(* IEC 61131-3 sources: SortJet_MasterSPS_Aufbau.fbsproj/09_Station/Stationen/Anlegetisch[201,205]/Aktionen, 2 files *)

(* ---- Anlegetisch_Austransport_FB_V01_00_00.fb.st ---- *)
(* METADATA
{
	"v3Meta": {
		"objectGuid": "29c6a30c-ea89-4d6e-bcb0-e2d154ff9fe9"
	}
}
*)
FUNCTION_BLOCK Anlegetisch_Austransport_FB_V01_00_00 EXTENDS Basic_Station_Austransport_FB_V01_00_00
(* Hinweis:
   - Austransport des Anlegetisches: Hubrahmen ausfahren, Austransport, Hubrahmen absenken, sobald die Sensorik
     frei ist, danach die Achsen des Glastransports abnullen
   - Der Rumpf ersetzt den Rumpf des Basic-Austransports, die Komponenten (Glastransport) kommen vom Basic-Baustein
*)
VAR_INPUT

  // Bausteine
  Hubrahmen : REFERENCE TO ZylinderPneumatik_Riemen_FB_V01_00_00;

END_VAR
//-------------------------------------------------------------------------------------------------
// AKTION: AUSTRANSPORT
//-------------------------------------------------------------------------------------------------
IF ( BasisStationsParameter.bAustransport[wWand]
     AND bpAutomatikAktiv )
THEN

  // Ausnahmesituation
  IF ( Glastransport.bpFehler ) THEN
    Glastransport.bpAustransport := FALSE;
    Glastransport.bpReferenz     := FALSE;
    BasisStationsParameter.wFehlerNummer := Glastransport.wpFehlerNr;
    steplAktion := STEP_900_E;
  END_IF

  IF ( Hubrahmen.bpFehler ) THEN
    Hubrahmen.bpStartAusfahren := FALSE;
    BasisStationsParameter.awFehlerInformationen[1] := cZYLINDER_HUBRAHMEN;
    BasisStationsParameter.wFehlerNummer := Hubrahmen.wpFehlerNr;
    steplAktion := STEP_900_E;
  END_IF

  CASE steplAktion OF
    // AUSTRANSPORT ==============================
    STEP_0_E:
      (* Hinweis:
         - -
      *)
      bpFehler := FALSE;
      Hubrahmen.bpStartAusfahren := NOT ( Hubrahmen.epStatusZylinder = eZylinderAusgefahren );

      steplAktion := STEP_10_E;

    // AUSTRANSPORT ==============================
    STEP_10_E:
      (* Anmerkung:
         - Hubpalette heben
      *)
      IF (  Hubrahmen.bpDone OR NOT Hubrahmen.bpStartAusfahren ) THEN
        Hubrahmen.bpStartAusfahren   := FALSE;
        Glastransport.bpAustransport := TRUE;
        steplAktion := STEP_30_E;
      END_IF

    // AUSTRANSPORT ==============================
    STEP_30_E:
      (* Hinweis:
         - Hubrahmen absenken wenn die Sensorik frei geworden ist
      *)
      IF Glastransport.bpSensorAuslauf THEN
        steplAktion := STEP_40_E;
      END_IF

      IF ( Glastransport.bpDone ) THEN
        Hubrahmen.bpStartEinfahren   := TRUE;
        Glastransport.bpAustransport := FALSE;
        steplAktion := STEP_50_E;
      END_IF

    // AUSTRANSPORT ==============================
    STEP_40_E:
      (* Hinweis:
         - Hubrahmen absenken wenn die Sensorik frei geworden ist
      *)
      IF (  NOT Glastransport.bpSensorAuslauf
           AND NOT BasisStationsParameter.InGlasTransportNachfolger[wWand].bEinlaufsensor )
      THEN
        Hubrahmen.bpStartEinfahren       := TRUE;
      END_IF

      IF ( Glastransport.bpDone ) THEN
        Hubrahmen.bpStartEinfahren       := TRUE;
        Glastransport.bpAustransport     := FALSE;
        steplAktion := STEP_50_E;
      END_IF

    // AUSTRANSPORT ==============================
    STEP_50_E:
      (* Hinweis:
         - Austransport ist vorbei: die Achsen des Glastransports abnullen (Zaehlerueberlauf des Gebers),
           nur nach dem Austransport, nie im Eintransport
      *)
      Glastransport.bpReferenz := TRUE;

      steplAktion := STEP_60_E;

    // AUSTRANSPORT ==============================
    STEP_60_E:
      IF ( Glastransport.bpDone ) THEN
        Glastransport.bpReferenz := FALSE;
        steplAktion := STEP_1000_E;
      END_IF

    // AUSTRANSPORT ==============================
    STEP_100_E:
      (* Anmerkung:
         - Hubpalette senken
      *)
      IF (  Hubrahmen.bpDone OR NOT BasisStationsParameter.stMKs.stStationsAufbau.bHubrahmen ) THEN
        Hubrahmen.bpStartEinfahren := FALSE;
        steplAktion := STEP_1000_E;
      END_IF

    // AUSTRANSPORT ==============================
    STEP_900_E:
      bpFehler := TRUE;
      BasisStationsParameter.bFehler := TRUE;
      BasisStationsParameter.bAustransportAbgeschlossen[wWand] := FALSE;

    // AUSTRANSPORT ==============================
    STEP_1000_E:
      BasisStationsParameter.bAustransportAbgeschlossen[wWand] := TRUE;

  // AUSTRANSPORT ==============================
  END_CASE
ELSE

  IF ( steplAktion > STEP_0_E ) THEN

    bpFehler := FALSE;
    Glastransport.bpAustransport := FALSE;
    Glastransport.bpReferenz     := FALSE;

    Hubrahmen.bpStartEinfahren := FALSE;
    Hubrahmen.bpStartAusfahren := FALSE;

    BasisStationsParameter.bAustransportAbgeschlossen[wWand] := FALSE;

    steplAktion := STEP_0_E;
  END_IF

END_IF
END_FUNCTION_BLOCK

(* ---- Anlegetisch_Eintransport_FB_V01_00_00.fb.st ---- *)
(* METADATA
{
	"v3Meta": {
		"objectGuid": "acd5983d-167d-4071-a6a9-aefc553f060d"
	}
}
*)
FUNCTION_BLOCK Anlegetisch_Eintransport_FB_V01_00_00 EXTENDS Basic_Station_Eintransport_FB_V01_00_00
(* Hinweis:
   - Eintransport des Anlegetisches von einer Fremdanlage (z.B. Brechanlage): Hubrahmen ausfahren, Anschlaege
     einfahren, Hoehenkontrolle positionieren, dann Eintransport
   - Mit dem Taster (oder wenn der Automatikbetrieb der Schneidlinie endet) wird die Scheibe nicht eintransportiert,
     sondern angelegt (bpAnlegenUmschalten)
   - Der Rumpf ersetzt den Rumpf des Basic-Eintransports, die Komponenten (Messachse, Glastransport) kommen vom Basic-Baustein
*)
VAR_INPUT

  // BOOLEAN
  bpAnlegenUmschalten : BOOL; // Station: Scheibe soll angelegt statt eintransportiert werden

  // Bausteine
  Anschlag  : REFERENCE TO ZylinderPneumatik_Anschlag_FB_V01_00_00;
  Hubrahmen : REFERENCE TO ZylinderPneumatik_Riemen_FB_V01_00_00;

END_VAR
VAR_OUTPUT

  // BOOLEAN
  bpAnlegenLampe : BOOL; // Ampel gruen / Signal Scheibe anlegen

END_VAR
//-------------------------------------------------------------------------------------------------
// AKTION: EINTRANSPORT
//-------------------------------------------------------------------------------------------------
IF( BasisStationsParameter.bEintransport[wWand]
    AND bpAutomatikAktiv )
THEN

  // Ausnahmesituation
  IF Hubrahmen.bpFehler THEN
    Hubrahmen.bpStartAusfahren := FALSE;
    BasisStationsParameter.awFehlerInformationen[1] := cZYLINDER_HUBRAHMEN;
    BasisStationsParameter.wFehlerNummer := Hubrahmen.wpFehlerNr;
    steplAktion := STEP_900_E;
  END_IF

  IF Anschlag.bpFehler THEN
    Anschlag.bpStartEinfahren := FALSE;
    BasisStationsParameter.awFehlerInformationen[1] := cZYLINDER_ANSCHLAG;
    BasisStationsParameter.wFehlerNummer := Anschlag.wpFehlerNr;
    steplAktion := STEP_900_E;
  END_IF

  IF Messachse.bpFehler THEN
    Messachse.bpPositionierung := FALSE;
    BasisStationsParameter.wFehlerNummer := Messachse.wpFehlerNr;
    steplAktion := STEP_900_E;
  END_IF

  CASE steplAktion OF
    // EINTRANSPORT ==================================
    STEP_0_E:

      bpFehler := FALSE;

      BasisStationsParameter.eStatusAuftrag   := eAuftragAktiv;

      IF ( bpGeblaeseFehler ) THEN
        BasisStationsParameter.wFehlerNummer := cMELDUNG_ANTRIEB_GEBLAESE;
        steplAktion := STEP_900_E;

      ELSE
        steplAktion := STEP_10_E;

      END_IF

    // EINTRANSPORT ==================================
    STEP_10_E:

      (* Anmerkung:
         - Glastransport Ausfahren
         - Anschläge einfahren
         - Messachse positionieren
      *)
      Hubrahmen.bpStartAusfahren := TRUE;
      Anschlag.bpStartEinfahren  := TRUE;

      IF Messachse.Antrieb.rpMaxPosition < ( BasisStationsParameter.pAuftrag[wWand].rAuftragsHoehe + Messachse.ppParameterBaustein.rKorrekturOffset ) THEN
        Messachse.rpZielPosition := Messachse.Antrieb.rpMaxPosition;
      ELSE
        Messachse.rpZielPosition := ( BasisStationsParameter.pAuftrag[wWand].rAuftragsHoehe + Messachse.ppParameterBaustein.rKorrekturOffset );
      END_IF
      Messachse.bpPositionierung := TRUE;

      steplAktion := STEP_20_E;

    // EINTRANSPORT ==================================
    STEP_20_E:

      (* Anmerkung:
         - Glastransport Ausfahren
         - Anschläge einfahren
         - Messachse.positionieren
      *)
      IF (     ( Hubrahmen.bpDone OR NOT BasisStationsParameter.stMKs.stStationsAufbau.bHubrahmen )
           AND Messachse.bpDone
           AND ( Anschlag.bpDone OR NOT BasisStationsParameter.stMKs.stStationsAufbau.bAnschlag ) )
      THEN
        Anschlag.bpStartEinfahren        := FALSE;
        Hubrahmen.bpStartAusfahren       := FALSE;
        Messachse.bpPositionierung := FALSE;
        steplAktion := STEP_30_E;
      END_IF

    // EINTRANSPORT ==================================
    STEP_30_E:

      (* Anmerkung:
         - Drosselklappe öffnen, damit auch sehr schweres Glas transportiert werden kann, indem die Luft das Glas leicht anhebt
      *)
      bpDrosselklappeOeffnen := TRUE;

      (* Anmerkung:
         - Glastransport Eintransport starten
      *)
      Glastransport.eGlastyp := BasisStationsParameter.wGlastyp[wWand];
      Glastransport.pAuftrag := BasisStationsParameter.pAuftrag[wWand];
      Glastransport.bpEintransport := TRUE;

      steplAktion := STEP_40_E;

      (* Fehlerbehandlung:
         - Glastransport
      *)
      IF Glastransport.bpFehler THEN
        Glastransport.bpEintransport := FALSE;
        BasisStationsParameter.wFehlerNummer := Glastransport.wpFehlerNr;
        steplAktion := STEP_900_E;
      END_IF

    // EINTRANSPORT ==================================
    STEP_40_E:

      bpAnlegenLampe  := TRUE;

      // Scheibe wird nicht Eintransportiert sondern soll angelegt werden
      IF bpAnlegenUmschalten THEN
        bpAnlegenLampe := FALSE;
        BasisStationsParameter.bAnlegen := TRUE;
        BasisStationsParameter.bEintransport[wWand] := FALSE;
      END_IF

      (* Anmerkung:
         - Auf den Glastransport warten
      *)
      IF Glastransport.bpDone THEN

        bpAnlegenLampe  := FALSE;

        Glastransport.bpEintransport := FALSE;
        BasisStationsParameter.eStatusAuftrag   := eAuftragErfolgreich;
        steplAktion := STEP_1000_E;
      END_IF

      (* Fehlerbehandlung:
         - Glastransport
         - Anschlag
      *)
      IF Glastransport.bpFehler THEN
        Glastransport.bpEintransport := FALSE;
        BasisStationsParameter.wFehlerNummer := Glastransport.wpFehlerNr;
        steplAktion := STEP_900_E;
      END_IF
      IF Anschlag.bpFehler THEN
        Anschlag.bpStartAusfahren := FALSE;
        BasisStationsParameter.awFehlerInformationen[1] := cZYLINDER_ANSCHLAG;
        BasisStationsParameter.wFehlerNummer := Anschlag.wpFehlerNr;
        steplAktion := STEP_900_E;
      END_IF

    // EINTRANSPORT ==================================
    STEP_900_E:
      bpFehler := TRUE;
      BasisStationsParameter.eStatusAuftrag   := eAuftragFehler;
      BasisStationsParameter.bFehler := TRUE;

    // EINTRANSPORT ==================================
    STEP_1000_E:
      BasisStationsParameter.dwWartezeit[wWand] := 0;
      BasisStationsParameter.bEintransportAbgeschlossen[wWand] := TRUE;

  // EINTRANSPORT ==================================
  END_CASE
ELSE

  IF( steplAktion > STEP_0_E )THEN
    bpFehler                              := FALSE;
    bpDrosselklappeOeffnen                := FALSE;
    Glastransport.bpEintransport          := FALSE;
    Anschlag.bpStartEinfahren             := FALSE;
    Anschlag.bpStartAusfahren             := FALSE;
    bpAnlegenLampe   := FALSE;
    Hubrahmen.bpStartAusfahren            := FALSE;
    Messachse.bpPositionierung      := FALSE;
    Messachse.bpVermessen_OberUndUnterkante_2_Sensoren := FALSE;
    BasisStationsParameter.bEintransportAbgeschlossen[wWand] := FALSE;
    steplAktion := STEP_0_E;
  END_IF

END_IF
END_FUNCTION_BLOCK
